Yaskawa INFORM job: 4043W1.JBI

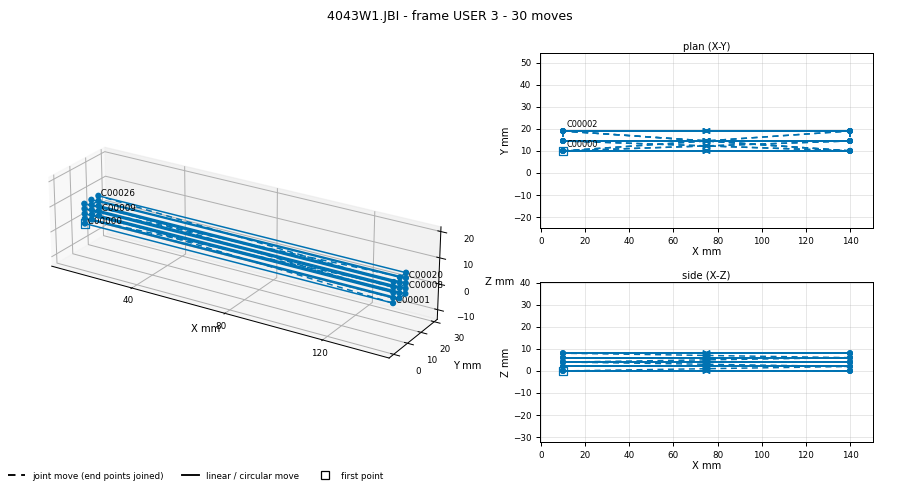
[picture p0: tool path of 4043W1.JBI in frame USER 3, 30 of 30 moves have a stored position in this frame; points joined in program order, loops and branches not executed]
/JOB
//NAME 4043W1
//POS
///NPOS 30,0,0,0,0,0
///USER 3
///TOOL 1
///POSTYPE USER
///RECTAN
///RCONF 1,0,0,0,0,0,0,0,0,0,0,0,0,0,0,0,0,0,0,0,0,0,0,0
C00000=10.000,10.000,0.000,0.0000,0.0000,-90.0000
C00001=140.000,10.000,0.000,0.0000,0.0000,-90.0000
C00002=10.000,19.000,0.000,0.0000,0.0000,-90.0000
C00003=140.000,19.000,0.000,0.0000,0.0000,-90.0000
C00004=140.000,14.500,0.000,0.0000,0.0000,-90.0000
C00005=10.000,14.500,0.000,0.0000,0.0000,-90.0000
C00006=140.000,10.000,2.000,0.0000,0.0000,-90.0000
C00007=10.000,10.000,2.000,0.0000,0.0000,-90.0000
C00008=140.000,19.000,2.000,0.0000,0.0000,-90.0000
C00009=10.000,19.000,2.000,0.0000,0.0000,-90.0000
C00010=10.000,14.500,2.000,0.0000,0.0000,-90.0000
C00011=140.000,14.500,2.000,0.0000,0.0000,-90.0000
C00012=10.000,10.000,4.000,0.0000,0.0000,-90.0000
C00013=140.000,10.000,4.000,0.0000,0.0000,-90.0000
C00014=10.000,19.000,4.000,0.0000,0.0000,-90.0000
C00015=140.000,19.000,4.000,0.0000,0.0000,-90.0000
C00016=140.000,14.500,4.000,0.0000,0.0000,-90.0000
C00017=10.000,14.500,4.000,0.0000,0.0000,-90.0000
C00018=140.000,10.000,6.000,0.0000,0.0000,-90.0000
C00019=10.000,10.000,6.000,0.0000,0.0000,-90.0000
C00020=140.000,19.000,6.000,0.0000,0.0000,-90.0000
C00021=10.000,19.000,6.000,0.0000,0.0000,-90.0000
C00022=10.000,14.500,6.000,0.0000,0.0000,-90.0000
C00023=140.000,14.500,6.000,0.0000,0.0000,-90.0000
C00024=10.000,10.000,8.000,0.0000,0.0000,-90.0000
C00025=140.000,10.000,8.000,0.0000,0.0000,-90.0000
C00026=10.000,19.000,8.000,0.0000,0.0000,-90.0000
C00027=140.000,19.000,8.000,0.0000,0.0000,-90.0000
C00028=140.000,14.500,8.000,0.0000,0.0000,-90.0000
C00029=10.000,14.500,8.000,0.0000,0.0000,-90.0000
//INST
///DATE 2025/03/17 13:38
///COMM Grasshopper
///ATTR SC,RW,RJ
////FRAME USER 3
///GROUP1 RB1
NOP
DOUT OT#(9) OFF
TIMER T=5.00
*LABEL0
MOVJ C00000 VJ=10.00 ACC=20
MACRO1 MJ#(0) ARGF202
ARCON
WVON WEV#(1)
MOVL C00001 V=10.0 ACC=20
WVOF
ARCOF
TIMER T=7.00
*LABEL1
MOVJ C00002 VJ=10.00 ACC=20
MACRO1 MJ#(0) ARGF202
ARCON
WVON WEV#(1)
MOVL C00003 V=10.0 ACC=20
WVOF
ARCOF
TIMER T=7.00
*LABEL2
MOVJ C00004 VJ=10.00 ACC=20
MACRO1 MJ#(0) ARGF202
ARCON
WVON WEV#(1)
MOVL C00005 V=10.0 ACC=20
WVOF
ARCOF
DOUT OT#(9) ON
TIMER T=70.00
DOUT OT#(9) OFF
TIMER T=13.00
*LABEL3
MOVJ C00006 VJ=10.00 ACC=20
MACRO1 MJ#(0) ARGF202
ARCON
WVON WEV#(1)
MOVL C00007 V=10.0 ACC=20
WVOF
ARCOF
TIMER T=7.00
*LABEL4
MOVJ C00008 VJ=10.00 ACC=20
MACRO1 MJ#(0) ARGF202
ARCON
WVON WEV#(1)
MOVL C00009 V=10.0 ACC=20
WVOF
ARCOF
TIMER T=7.00
*LABEL5
MOVJ C00010 VJ=10.00 ACC=20
MACRO1 MJ#(0) ARGF202
ARCON
WVON WEV#(1)
MOVL C00011 V=10.0 ACC=20
WVOF
ARCOF
DOUT OT#(9) ON
TIMER T=70.00
DOUT OT#(9) OFF
TIMER T=13.00
*LABEL6
MOVJ C00012 VJ=10.00 ACC=20
MACRO1 MJ#(0) ARGF202
ARCON
WVON WEV#(1)
MOVL C00013 V=10.0 ACC=20
WVOF
ARCOF
TIMER T=7.00
*LABEL7
MOVJ C00014 VJ=10.00 ACC=20
MACRO1 MJ#(0) ARGF202
ARCON
WVON WEV#(1)
MOVL C00015 V=10.0 ACC=20
WVOF
ARCOF
TIMER T=7.00
*LABEL8
MOVJ C00016 VJ=10.00 ACC=20
MACRO1 MJ#(0) ARGF202
ARCON
WVON WEV#(1)
MOVL C00017 V=10.0 ACC=20
WVOF
ARCOF
DOUT OT#(9) ON
TIMER T=70.00
DOUT OT#(9) OFF
TIMER T=13.00
*LABEL9
MOVJ C00018 VJ=10.00 ACC=20
MACRO1 MJ#(0) ARGF202
ARCON
WVON WEV#(1)
MOVL C00019 V=10.0 ACC=20
WVOF
ARCOF
TIMER T=7.00
*LABEL10
MOVJ C00020 VJ=10.00 ACC=20
MACRO1 MJ#(0) ARGF202
ARCON
WVON WEV#(1)
MOVL C00021 V=10.0 ACC=20
WVOF
ARCOF
TIMER T=7.00
*LABEL11
MOVJ C00022 VJ=10.00 ACC=20
MACRO1 MJ#(0) ARGF202
ARCON
WVON WEV#(1)
MOVL C00023 V=10.0 ACC=20
WVOF
ARCOF
DOUT OT#(9) ON
TIMER T=70.00
DOUT OT#(9) OFF
TIMER T=13.00
*LABEL12
MOVJ C00024 VJ=10.00 ACC=20
MACRO1 MJ#(0) ARGF202
ARCON
WVON WEV#(1)
MOVL C00025 V=10.0 ACC=20
WVOF
ARCOF
TIMER T=7.00
*LABEL13
MOVJ C00026 VJ=10.00 ACC=20
MACRO1 MJ#(0) ARGF202
ARCON
WVON WEV#(1)
MOVL C00027 V=10.0 ACC=20
WVOF
ARCOF
TIMER T=7.00
*LABEL14
MOVJ C00028 VJ=10.00 ACC=20
MACRO1 MJ#(0) ARGF202
ARCON
WVON WEV#(1)
MOVL C00029 V=10.0 ACC=20
WVOF
ARCOF
DOUT OT#(9) ON
TIMER T=70.00
DOUT OT#(9) OFF
TIMER T=13.00
END
